FUNCTION_BLOCK PRINT_QUEUE
  {SET_ATTRIBUTE(OpcUa, SERVICE)}
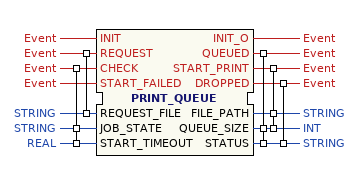
  EVENT_INPUT
    INIT;
    REQUEST WITH REQUEST_FILE;
    CHECK WITH JOB_STATE, START_TIMEOUT;
    START_FAILED;
  END_EVENT
  EVENT_OUTPUT
    INIT_O;
    QUEUED WITH QUEUE_SIZE, STATUS;
    START_PRINT WITH FILE_PATH, QUEUE_SIZE;
    DROPPED WITH STATUS;
  END_EVENT
  VAR_INPUT
    REQUEST_FILE : STRING; {SET_ATTRIBUTE(OpcUa, Variable)}
    JOB_STATE : STRING; {SET_ATTRIBUTE(OpcUa, Variable)}
    START_TIMEOUT : REAL; {SET_ATTRIBUTE(OpcUa, Constant)}
  END_VAR
  VAR_OUTPUT
    FILE_PATH : STRING; {SET_ATTRIBUTE(OpcUa, Variable)}
    QUEUE_SIZE : INT; {SET_ATTRIBUTE(OpcUa, Variable)}
    STATUS : STRING; {SET_ATTRIBUTE(OpcUa, Variable)}
  END_VAR
END_FUNCTION_BLOCK
